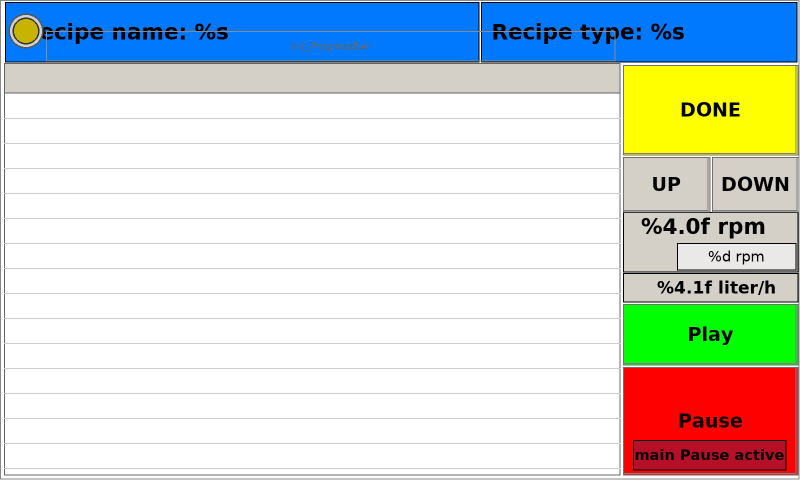
VISUALIZATION vis_Dissolve  // 800x480
VAR_IN_OUT
	
END_VAR

VAR
	lacal_bool: BOOL:=TRUE;
END_VAR
    Table (4,63 616x412), data array: stPLC_To_VisuPLC.arr_Component
        p3854506369: stPLC_To_VisuPLC.arr_Component[INDEX].sDescription
        p1892666644: stPLC_To_VisuPLC.arr_Component[INDEX].eIngredientType
        p338671338: stPLC_To_VisuPLC.arr_Component[INDEX].rWeight
        p2170511999: stPLC_To_VisuPLC.arr_Component[INDEX].rWeightPercentage
        p3723444502: stPLC_To_VisuPLC.arr_Component[INDEX].rFlowRate_Dissolving
        p1218418051: stPLC_To_VisuPLC.arr_Component[INDEX].rFlowRate_Blending
        p746581629: stPLC_To_VisuPLC.arr_Component[INDEX].tBlendingDuration
        p2232123230: Component Description
        p1755163831: Weight [kg]
        p4092479075: %
        p2237128397: Flow [RPM]
        p1137915858: stPLC_To_VisuPLC.iActual_Component
    Rectangle (623,212 175x60), "%4.0f rpm", text variable: g_HMI_Panel.stVisuPLC_To_PLC.RPM_setPoint
    Button (623,157 87x55), "UP", input disabled if: NOT g_HMI_Panel.stPLC_To_VisuPLC.bDissolving_Active
        OnMouseDown: execute {
            g_HMI_Panel.stVisuPLC_To_PLC.RPM_setPoint:=
            g_HMI_Panel.stVisuPLC_To_PLC.RPM_setPoint+50;
            IF g_HMI_Panel.stVisuPLC_To_PLC.RPM_setPoint>2500 THEN;
            	g_HMI_Panel.stVisuPLC_To_PLC.RPM_setPoint:=2500;
            END_IF
        }
    Button (712,157 87x55), "DOWN", input disabled if: NOT g_HMI_Panel.stPLC_To_VisuPLC.bDissolving_Active
        OnMouseDown: execute {
            g_HMI_Panel.stVisuPLC_To_PLC.RPM_setPoint:=
            g_HMI_Panel.stVisuPLC_To_PLC.RPM_setPoint-50;
            IF g_HMI_Panel.stVisuPLC_To_PLC.RPM_setPoint<300 THEN;
            	g_HMI_Panel.stVisuPLC_To_PLC.RPM_setPoint:=300;
            END_IF
        }
    Rectangle (5,2 474x60), "Recipe name: %s", text variable: g_HMI_Panel.stPLC_To_VisuPLC.Description
    Lamp1 (6,11 40x40), variable: g_HMI_Panel.stPLC_To_VisuPLC.lifeBit, style: Lamp-Lamp1-Yellow
    Rectangle (677,243 119x27), "%d rpm", text variable: g_HMI_Panel.stPLC_To_VisuPLC.RPM_FeedBack
    Rectangle (481,2 316x60), "Recipe type: %s", text variable: g_HMI_Panel.stPLC_To_VisuPLC.prodType
    Button (623,367 175x108), "Pause", colour toggle: g_HMI_Panel.stVisuPLC_To_PLC.bPauseTriBlender, pressed state: g_HMI_Panel.stVisuPLC_To_PLC.bPauseTriBlender, input disabled if: g_HMI_Panel.stVisuPLC_To_PLC.bPauseTriBlender OR NOT g_HMI_Panel.stPLC_To_VisuPLC.bDissolving_Active
        toggle g_HMI_Panel.stVisuPLC_To_PLC.bPauseTriBlender
    Button (623,304 175x61), "Play", colour toggle: NOT g_HMI_Panel.stVisuPLC_To_PLC.bPauseTriBlender, pressed state: NOT g_HMI_Panel.stVisuPLC_To_PLC.bPauseTriBlender, input disabled if: NOT g_HMI_Panel.stVisuPLC_To_PLC.bPauseTriBlender
        toggle g_HMI_Panel.stVisuPLC_To_PLC.bPauseTriBlender
    Button (623,65 175x90), "DONE", input disabled if: NOT g_HMI_Panel.stPLC_To_VisuPLC.bDissolving_Active OR g_HMI_Panel.stVisuPLC_To_PLC.bPauseTriBlender
        OnMouseClick: execute { g_HMI_Panel.stVisuPLC_To_PLC.bActualComponentDisolving_Done:=TRUE; }
    Rectangle (3,100 618x378)
    Frame (46,31 569x30), invisible if: NOT g_HMI_Panel.stPLC_To_VisuPLC.bBlending_Active
        shows vis_ProgressBar()
        p2738717112: MAIN.iProgressBarOfset
    Rectangle (623,273 175x29), "%4.1f liter/h", text variable: g_HMI_Panel.stPLC_To_VisuPLC.Flow_FeedBack
    Rectangle (633,440 153x30), "main Pause active", invisible if: NOT g_HMI_Panel.stPLC_To_VisuPLC.bMainPause_Active
END_VISUALIZATION

(* stored: Version 1.1.0.1, ProductVersion 3.1.4024.15
   Visu vis_Dissolve: Id {919e275f-691e-4ef6-b817-488a1cc80f7e} *)
